(* IEC 61131-3 sources: Test-Git_ESME26/TestProgettoESME_26.fbsproj/AxisModule_Migration_Example.device.xml.v3^/Plc Logic.plclogic.xml.v3^/Application.application.xml.v3^/Test_AxisModule, 2 files *)

(* ---- Global_ExceptionList.gvl ---- *)
VAR_GLOBAL
		(* ExceptionHandling and Logging *)
	G_stExceptionList			: TPL.ST_ExceptionList;
	G_stLogDataList				: TPL.ST_LogDataList;

END_VAR

(* ---- GVL_Encoder.gvl ---- *)
VAR_GLOBAL
	LE_Master		: MOIN.FB_LogicalEncoder;
	LE_Slave1		: MOIN.FB_LogicalEncoder;
	LE_Slave2		: MOIN.FB_LogicalEncoder;
END_VAR
